(*
SPDX-FileCopyrightText: © 2026 Oleksandr Tiutyk <trofimich@gmail.com>
SPDX-License-Identifier: MIT
License: https://opensource.org/license/mit
*)

(*!
<summary>Provides fluent assertions on a copied WSTRING(255) value.</summary>
<description>
Copies actual into persistent instance storage before the entry method returns; literals and expression
results therefore remain valid throughout the immediate chain. Owns no heap allocation or pointed-to resource.
The message prefixes every failure until the next preparation. Finish one chain before starting another on
the owning Assertions provider. Use only from the owning test callback on one task, without reentry.
Obtain this context from the owning provider; direct unprepared use is unsupported.
Expected arguments use the declared IEC type; ordinary compiler conversions happen before comparison.
This context does not depend on another assertion context.
Object metadata is available before preparation; inherited equality compares instance identity.
Actual and expected strings are limited to 255 characters; normal IEC parameter conversion may truncate
longer inputs. Use the generic That entry with live variables for longer strings. Comparison is by code unit.
</description>
*)

{attribute 'no_explicit_call' := 'do not call this function block directly'}
FUNCTION_BLOCK WideStringAssertionContext EXTENDS TOF_Core.Object
VAR_STAT
	{attribute 'hide'}
	_ClassName : STRING := __POUNAME();
END_VAR
VAR
	_Actual : WSTRING(255);
	_TestCase : ITestCase;
	_Message : WSTRING(255);
END_VAR

(*!
<summary>Provides the implementation class name.</summary>
<description>
Borrowed read-only reference to compiler-initialized storage, valid throughout the instance lifetime.
Do not modify the returned reference; no ownership is transferred.
</description>
*)
{attribute 'monitoring' := 'call'}
PROPERTY ClassName : REFERENCE TO STRING
GET
ClassName REF= _ClassName;
END_GET
END_PROPERTY

(*!
<summary>Asserts that the actual value is strictly greater than expected.</summary>
<description>
Records failure without interrupting the callback; preserves the message for the rest of the chain.
</description>
<param name="expected">Expected value converted by the compiler to WSTRING(255).</param>
*)
METHOD FINAL IsGreaterThan : REFERENCE TO WideStringAssertionContext
VAR_INPUT
	expected : WSTRING(255);
END_VAR
VAR
	comparison : TOF_Core.COMPARISON_RESULT;
END_VAR
comparison := compareExpected(expected := expected);

IF comparison <> TOF_Core.COMPARISON_RESULT.FIRST_GREATER_THAN_SECOND THEN
	failComparison(
		expected := expected,
		expectation := "Expected value > "
	);
END_IF

IsGreaterThan REF= THIS^;
END_METHOD

(*!
<summary>Asserts that the actual value meets the inclusive lower boundary.</summary>
<description>
Records failure without interrupting the callback; preserves the message for the rest of the chain.
</description>
<param name="expected">Expected value converted by the compiler to WSTRING(255).</param>
*)
METHOD FINAL IsGreaterThanOrEquals : REFERENCE TO WideStringAssertionContext
VAR_INPUT
	expected : WSTRING(255);
END_VAR
VAR
	comparison : TOF_Core.COMPARISON_RESULT;
END_VAR
comparison := compareExpected(expected := expected);

IF comparison = TOF_Core.COMPARISON_RESULT.FIRST_LESS_THAN_SECOND THEN
	failComparison(
		expected := expected,
		expectation := "Expected value >= "
	);
END_IF

IsGreaterThanOrEquals REF= THIS^;
END_METHOD

(*!
<summary>Asserts that the actual value is strictly less than expected.</summary>
<description>
Records failure without interrupting the callback; preserves the message for the rest of the chain.
</description>
<param name="expected">Expected value converted by the compiler to WSTRING(255).</param>
*)
METHOD FINAL IsLessThan : REFERENCE TO WideStringAssertionContext
VAR_INPUT
	expected : WSTRING(255);
END_VAR
VAR
	comparison : TOF_Core.COMPARISON_RESULT;
END_VAR
comparison := compareExpected(expected := expected);

IF comparison <> TOF_Core.COMPARISON_RESULT.FIRST_LESS_THAN_SECOND THEN
	failComparison(
		expected := expected,
		expectation := "Expected value < "
	);
END_IF

IsLessThan REF= THIS^;
END_METHOD

(*!
<summary>Asserts that the actual value meets the inclusive upper boundary.</summary>
<description>
Records failure without interrupting the callback; preserves the message for the rest of the chain.
</description>
<param name="expected">Expected value converted by the compiler to WSTRING(255).</param>
*)
METHOD FINAL IsLessThanOrEquals : REFERENCE TO WideStringAssertionContext
VAR_INPUT
	expected : WSTRING(255);
END_VAR
VAR
	comparison : TOF_Core.COMPARISON_RESULT;
END_VAR
comparison := compareExpected(expected := expected);

IF comparison = TOF_Core.COMPARISON_RESULT.FIRST_GREATER_THAN_SECOND THEN
	failComparison(
		expected := expected,
		expectation := "Expected value <= "
	);
END_IF

IsLessThanOrEquals REF= THIS^;
END_METHOD

(*!
<summary>Provides the library namespace.</summary>
<description>
Borrowed read-only reference to the compiler-initialized namespace, valid throughout the instance lifetime.
Do not modify the returned reference; no ownership is transferred.
</description>
*)
{attribute 'monitoring' := 'call'}
PROPERTY NamespaceName : REFERENCE TO STRING
GET
NamespaceName REF= CurrentNamespace.Name;
END_GET
END_PROPERTY

(*!
<summary>Asserts inequality with the expected value.</summary>
<description>
Records failure without interrupting the callback; preserves the message for the rest of the chain.
</description>
<param name="expected">Expected value converted by the compiler to WSTRING(255).</param>
*)
METHOD FINAL NotToBe : REFERENCE TO WideStringAssertionContext
VAR_INPUT
	expected : WSTRING(255);
END_VAR
VAR
	comparison : TOF_Core.COMPARISON_RESULT;
END_VAR
comparison := compareExpected(expected := expected);

IF comparison = TOF_Core.COMPARISON_RESULT.FIRST_EQUAL_TO_SECOND THEN
	failComparison(
		expected := expected,
		expectation := "Expected value not to be: "
	);
END_IF

NotToBe REF= THIS^;
END_METHOD

(*!
<summary>Copies the actual operand and replaces the chain-wide message.</summary>
<description>
Called by the owning Assertions provider after it verifies the running test case.
No pointer to this method's input storage is retained. The receiver is borrowed until the next preparation;
the owning provider keeps it alive throughout the immediate chain.
</description>
<param name="actual">Value copied into this context.</param>
<param name="testCase">Borrowed failure receiver for the immediate chain.</param>
<param name="message">Copied diagnostic prefix, including empty to clear the previous prefix.</param>
*)
METHOD INTERNAL FINAL Prepare
VAR_INPUT
	actual : WSTRING(255);
	testCase : ITestCase;
	message : WSTRING(255);
END_VAR
_Actual := actual;
_TestCase := testCase;
_Message := message;
END_METHOD

(*!
<summary>Reports the byte size of this concrete instance.</summary>
<description>
Includes inline fields and nested instances, but excludes separately allocated payloads.
Obtaining the size does not transfer ownership or validate an arbitrary address.
</description>
*)
{attribute 'monitoring' := 'call'}
PROPERTY SelfSize : ULINT
GET
SelfSize := XSIZEOF(THIS^);
END_GET
END_PROPERTY

(*!
<summary>Asserts equality with the expected value.</summary>
<description>
Records failure without interrupting the callback; preserves the message for the rest of the chain.
</description>
<param name="expected">Expected value converted by the compiler to WSTRING(255).</param>
*)
METHOD FINAL ToBe : REFERENCE TO WideStringAssertionContext
VAR_INPUT
	expected : WSTRING(255);
END_VAR
VAR
	comparison : TOF_Core.COMPARISON_RESULT;
END_VAR
comparison := compareExpected(expected := expected);

IF comparison <> TOF_Core.COMPARISON_RESULT.FIRST_EQUAL_TO_SECOND THEN
	failComparison(
		expected := expected,
		expectation := "Expected: "
	);
END_IF

ToBe REF= THIS^;
END_METHOD

(*!
<summary>Asserts that the copied string contains the specified substring.</summary>
<description>
Uses the context's string encoding and retains the chain message after the assertion.
</description>
<param name="substring">Substring of at most 255 characters in the same encoding.</param>
*)
METHOD FINAL ToContain : REFERENCE TO WideStringAssertionContext
VAR_INPUT
	substring : WSTRING(255);
END_VAR
VAR
	actualText : WSTRING(255);
	expectedText : WSTRING(255);
	diagnostic : TOF_Core.ERROR_MESSAGE;
END_VAR
IF NOT TOF_Core.WideStrings.Contains(stringToSearchIn := _Actual, stringToFind := substring) THEN
	actualText := _Actual;
	expectedText := substring;

	diagnostic := TOF_Core.WideStrings.Concat255(
		"Expected text to contain '",
		expectedText,
		"', but was: '",
		actualText,
		"'"
	);

	TestServices.ReportAssertionFailure(
		testCase := _TestCase,
		message := _Message,
		sourceClassName := ClassName,
		defaultMessage := diagnostic
	);
END_IF

ToContain REF= THIS^;
END_METHOD

(*!
<summary>Compares the copied string with a typed boundary by code unit.</summary>
<description>
Both typed operands provide terminated storage. Reads through the first differing code unit or
terminator; does not allocate, convert encodings or retain the expected storage.
</description>
<param name="expected">Same-encoding boundary alive for this call.</param>
*)
METHOD PRIVATE compareExpected : TOF_Core.COMPARISON_RESULT
VAR_INPUT
	expected : WSTRING(255);
END_VAR
VAR
	actualData : POINTER TO WORD;
	expectedData : POINTER TO WORD;
	characterIndex : UDINT;
END_VAR
actualData := ADR(_Actual);
expectedData := ADR(expected);

WHILE TRUE DO
	IF actualData[characterIndex] < expectedData[characterIndex] THEN
		compareExpected := TOF_Core.COMPARISON_RESULT.FIRST_LESS_THAN_SECOND;
		RETURN;
	ELSIF actualData[characterIndex] > expectedData[characterIndex] THEN
		compareExpected := TOF_Core.COMPARISON_RESULT.FIRST_GREATER_THAN_SECOND;
		RETURN;
	ELSIF actualData[characterIndex] = TO_WORD(TOF_Core.UnsignedInt16.MIN_VALUE) THEN
		compareExpected := TOF_Core.COMPARISON_RESULT.FIRST_EQUAL_TO_SECOND;
		RETURN;
	END_IF

	characterIndex := characterIndex + 1;
END_WHILE
END_METHOD

(*!
<summary>Formats a failed typed predicate and reports it with the chain message.</summary>
<description>
Does not change operands or chain state. The receiver retains its first failure. Reporting exceptions
propagate to the enclosing test callback handler; an unprepared receiver is a configuration error.
</description>
<param name="expected">Typed expected operand used only for this diagnostic.</param>
<param name="expectation">Prefix identifying the failed predicate.</param>
*)
METHOD PRIVATE failComparison
VAR_INPUT
	expected : WSTRING(255);
	expectation : WSTRING(40);
END_VAR
VAR
	actualText : WSTRING(255);
	expectedText : WSTRING(255);
	diagnostic : TOF_Core.ERROR_MESSAGE;
END_VAR
actualText := _Actual;
expectedText := expected;

diagnostic := TOF_Core.WideStrings.Concat255(
	expectation,
	expectedText,
	", but was: ",
	actualText
);

TestServices.ReportAssertionFailure(
	testCase := _TestCase,
	message := _Message,
	sourceClassName := ClassName,
	defaultMessage := diagnostic
);
END_METHOD

END_FUNCTION_BLOCK

(* stored: Version 1.1.0.1
   POU WideStringAssertionContext: Id {bd0d153b-0cfe-48b0-beb1-1dcf91d1c22f}, SpecialFunc None
   Folder Service methods: Id {393cb245-ba1c-4c91-9698-d88546433a30}
   Property ClassName: Id {1d3edba2-ace0-4287-b14b-4694456b05a0}
   Get Get: Id {10225fec-44d2-4fa9-b1b8-17c22abe5b6b}
   Method IsGreaterThan: Id {4a6ae0c9-db85-4c5d-9c5f-acd126653b88}
   Method IsGreaterThanOrEquals: Id {24b95cc1-bca1-4f9a-85e7-93d782b3df6f}
   Method IsLessThan: Id {3ca1221a-1172-4da3-a5d8-e119e8942d18}
   Method IsLessThanOrEquals: Id {3573d853-e0d8-44fc-9f01-9c3e316e2d48}
   Property NamespaceName: Id {79419c8c-6ccc-435e-be34-5dce5d62accb}
   Get Get: Id {6325c5ff-6c92-414c-a3f2-6cae0b6667ba}
   Method NotToBe: Id {afb59a13-41f0-461f-a865-7b555e017df2}
   Method Prepare: Id {4a5fb132-3682-4f7a-b1e5-e5cdd9d6dd7a}
   Property SelfSize: Id {940e583e-d3c2-415d-8a32-349f469c8fdd}
   Get Get: Id {4268546e-1b7f-476d-bbed-fcfd5bde8a55}
   Method ToBe: Id {8723f87b-2a45-4eba-9930-c4e4578fe18c}
   Method ToContain: Id {6acb9c6e-c24a-434d-956d-47f1edbd34fd}
   Method compareExpected: Id {118f1099-9db8-403d-84d4-9e18a40e984c}
   Method failComparison: Id {3637e56c-4414-4f1a-a8e6-44a959e8618a} *)
